(* IEC 61131-3 sources: repolevel_ST_code_completion/output/full_case_fixed/repoeval_plc_hello_mixing_tank/readful_result, 1 file *)

(* ---- FB_AutoSequence.st ---- *)
FUNCTION_BLOCK FB_AutoSequence
VAR_INPUT
	bEnable				:	BOOL;			// 使能自动序列
	bReset				:	BOOL;			// 复位到排空状态

	// 液位传感器反馈
	bTankLevelFull		:	BOOL;			// 液位满传感器
	bTankLevelEmpty		:	BOOL;			// 液位空传感器

	// 设备状态反馈
	bMixerRunning		:	BOOL;			// 混合电机运行中
	bMedium1Opened		:	BOOL;			// 介质1阀门打开
	bMedium2Opened		:	BOOL;			// 介质2阀门打开
	bDrainOpened		:	BOOL;			// 排空阀门打开

	// 配置参数
	tMixingDuration		:	TIME := T#10S;	// 混合持续时间
END_VAR
VAR_OUTPUT
	// 设备控制输出
	bMixerRunCmd		:	BOOL;			// 混合电机运行命令
	bMedium1OpenCmd		:	BOOL;			// 介质1阀门打开命令
	bMedium2OpenCmd		:	BOOL;			// 介质2阀门打开命令
	bDrainOpenCmd		:	BOOL;			// 排空阀门打开命令

	// 状态输出
	eCurrentState		:	AUTO_SEQUENCE;	// 当前状态
	nCyclesCompleted	:	UINT;			// 完成的循环次数
END_VAR
VAR
	tonMixing			:	TON;			// 混合定时器
END_VAR

// Reset logic
IF bReset THEN
	eCurrentState := AUTO_SEQUENCE.DRAINING;
	nCyclesCompleted := 0;
END_IF

// Automatic sequence state machine
IF bEnable THEN
	CASE eCurrentState OF
		AUTO_SEQUENCE.FILLING:
			// Ensure other devices are not operating
			bMixerRunCmd := FALSE;
			bDrainOpenCmd := FALSE;

			// Open medium valves to fill the tank
			bMedium1OpenCmd := TRUE;
			bMedium2OpenCmd := TRUE;

			// Transition to mixing state when tank is full
			IF bTankLevelFull THEN
				eCurrentState := AUTO_SEQUENCE.MIXING;
			END_IF;

		AUTO_SEQUENCE.MIXING:
			// Ensure filling and draining are stopped
			bMedium1OpenCmd := FALSE;
			bMedium2OpenCmd := FALSE;
			bDrainOpenCmd := FALSE;

			// Start mixer
			bMixerRunCmd := TRUE;

			// Activate mixing timer
			tonMixing(IN := TRUE, PT := tMixingDuration);

			// Transition to draining state when mixing is complete
			IF tonMixing.Q THEN
				eCurrentState := AUTO_SEQUENCE.DRAINING;
			END_IF;

		AUTO_SEQUENCE.DRAINING:
			// Ensure filling and mixing are stopped
			bMedium1OpenCmd := FALSE;
			bMedium2OpenCmd := FALSE;
			bMixerRunCmd := FALSE;

			// Open drain valve to empty the tank
			bDrainOpenCmd := TRUE;

			// Transition to filling state when tank is empty
			IF bTankLevelEmpty THEN
				eCurrentState := AUTO_SEQUENCE.FILLING;
				nCyclesCompleted := nCyclesCompleted + 1;
			END_IF;

		// Default case to handle unexpected states
		ELSE
			// Reset all commands
			bMixerRunCmd := FALSE;
			bMedium1OpenCmd := FALSE;
			bMedium2OpenCmd := FALSE;
			bDrainOpenCmd := FALSE;

			// Transition to draining state
			eCurrentState := AUTO_SEQUENCE.DRAINING;
	END_CASE;
END_IF;
END_FUNCTION_BLOCK
